TYPE E_OperationButtons :(
	ePauseAll:=0,
	ePlayAll:=1);
END_TYPE

(* stored: Version 1.1.0.1, ProductVersion 3.1.4024.13
   DUT E_OperationButtons: Id {9b040a80-05b8-49a9-89be-4993401fa1e7} *)
